// TIA Portal V21 export
// export: Created 2026-10-25T15:00:20.9672797Z, ExportSetting WithDefaults, DisplayName Totally Integrated Automation Portal, DisplayVersion V21 Update 3, DisplayName TIA Portal Test Suite Advanced, DisplayVersion V21 Update 1, DisplayName SINAMICS Startdrive Advanced, DisplayVersion V21 Update 1, DisplayName SINAMICS Startdrive G130, G150, S120, S150, G200, G210, G210C, G210X, G220, S200, S210, S220, Innomotics MVD, DisplayVersion V21 Update 1, DisplayName SINAMICS Startdrive G110M, G120, G120C, G120D, G120P, G115D, DisplayVersion V21 Update 1, DisplayName STEP 7 Professional, DisplayVersion V21 Update 3, DisplayName STEP 7 Safety, DisplayVersion V21, DisplayName Tech WebApplication, DisplayVersion V21, DisplayName WinCC Basic/Comfort/Advanced, DisplayVersion V21 Update 3, DisplayName WinCC Professional, DisplayVersion V21 Update 3, DisplayName WinCC Unified, DisplayVersion V21 Update 3
FUNCTION_BLOCK "TgpNamespace_NumericFC_LAD"   // FB5, LAD
VERSION : 0.1
// stored: Access Unpublished, AutoNumber true, IsIECCheckEnabled false, IsRetainMemResEnabled false, MemoryReserve 100, Namespace TiaMcp_UnitA.Alternate, SetENOAutomatically false, UDAEnableTagReadback false
   VAR_INPUT
      Value : Int;
   END_VAR
   VAR_OUTPUT
      Result : Int;
      Returned : Int;
   END_VAR
   VAR_IN_OUT
      Accumulator : Int;
   END_VAR
BEGIN

REGION Network 1
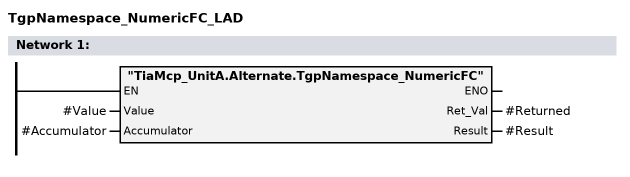
   RUNG wire#powerrail
      "TiaMcp_UnitA.Alternate.TgpNamespace_NumericFC"(Value := #Value, Accumulator := #Accumulator, Result => #Result, Ret_Val => #Returned)
   END_RUNG
   // the same network as SCL:
   #Returned := "TiaMcp_UnitA.Alternate.TgpNamespace_NumericFC"(Value := #Value,
                           Accumulator := #Accumulator,
                           Result => #Result);
END_REGION
END_FUNCTION_BLOCK
